// TIA Portal V17 export
// export: Created 2026-11-08T05:50:28.6935429Z, ExportSetting WithDefaults, DisplayName Totally Integrated Automation Portal, DisplayVersion V17, DisplayName TIA Portal Openness, DisplayVersion V17, DisplayName TIA Portal Version Control Interface, DisplayVersion V17, DisplayName STEP 7 Professional, DisplayVersion V17, DisplayName STEP 7 Safety, DisplayVersion V17, DisplayName WinCC Professional, DisplayVersion V17
FUNCTION_BLOCK "FB_Motor_Banderas"   // FB3, LAD
TITLE = Arranque y paro por BANDERAS (S/R)
{ S7_Optimized_Access := 'TRUE' }
VERSION : 0.1
// Estilo clásico: bandera de marcha con SET/RESET (paro dominante). Sin térmico se para; al recuperarse el térmico se puede volver a arrancar sin RESET.
// stored: AutoNumber true, IsIECCheckEnabled false, IsRetainMemResEnabled false, MemoryReserve 100, SetENOAutomatically false, UDAEnableTagReadback false
   VAR_INPUT
      Marcha : Bool;   // Orden de marcha (pulsador o HMI)
      Paro : Bool;   // Orden de paro: 1 = parar
      Termico_OK : Bool;   // 1 = relé térmico sin falla
      Reset : Bool;   // Reset de falla
   END_VAR
   VAR_OUTPUT
      Motor : Bool;   // Orden al contactor
      Piloto_Marcha : Bool;   // Piloto verde
      Piloto_Falla : Bool;   // Piloto rojo
      Estado : Int;   // 0 Reposo, 10 Marcha, 90 Falla
   END_VAR
   VAR
      B_Marcha : Bool;   // Bandera: motor en marcha
      B_Falla : Bool;   // Bandera: falla térmico
   END_VAR
BEGIN

REGION Network 1: SET bandera de marcha
   // Marcha sin paro y con térmico OK.
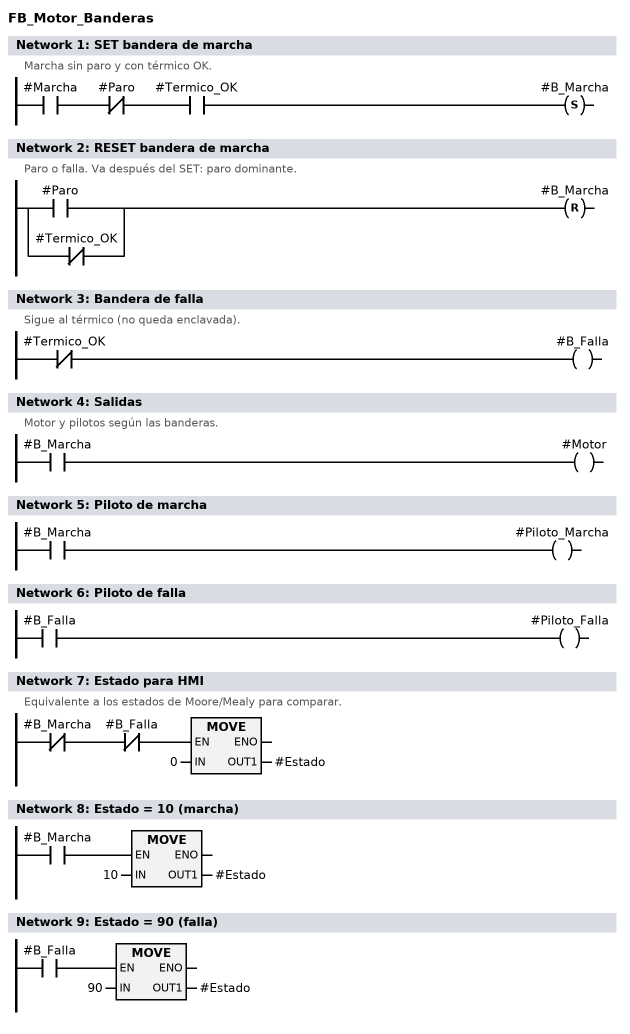
   RUNG wire#powerrail
      Contact( #Marcha )
      I_Contact( #Paro )
      Contact( #Termico_OK )
      S_Coil( #B_Marcha )
   END_RUNG
   // the same network as SCL:
   IF #Marcha AND NOT #Paro AND #Termico_OK THEN #B_Marcha := TRUE; END_IF;
END_REGION

REGION Network 2: RESET bandera de marcha
   // Paro o falla. Va después del SET: paro dominante.
   RUNG wire#powerrail
      Contact( #Paro )
      wire#w1
      R_Coil( #B_Marcha )
   END_RUNG
   RUNG wire#powerrail
      I_Contact( #Termico_OK )
   END_RUNG wire#w1
   // the same network as SCL:
   IF #Paro OR NOT #Termico_OK THEN #B_Marcha := FALSE; END_IF;
END_REGION

REGION Network 3: Bandera de falla
   // Sigue al térmico (no queda enclavada).
   RUNG wire#powerrail
      I_Contact( #Termico_OK )
      Coil( #B_Falla )
   END_RUNG
   // the same network as SCL:
   #B_Falla := NOT #Termico_OK;
END_REGION

REGION Network 4: Salidas
   // Motor y pilotos según las banderas.
   RUNG wire#powerrail
      Contact( #B_Marcha )
      Coil( #Motor )
   END_RUNG
   // the same network as SCL:
   #Motor := #B_Marcha;
END_REGION

REGION Network 5: Piloto de marcha
   RUNG wire#powerrail
      Contact( #B_Marcha )
      Coil( #Piloto_Marcha )
   END_RUNG
   // the same network as SCL:
   #Piloto_Marcha := #B_Marcha;
END_REGION

REGION Network 6: Piloto de falla
   RUNG wire#powerrail
      Contact( #B_Falla )
      Coil( #Piloto_Falla )
   END_RUNG
   // the same network as SCL:
   #Piloto_Falla := #B_Falla;
END_REGION

REGION Network 7: Estado para HMI
   // Equivalente a los estados de Moore/Mealy para comparar.
   RUNG wire#powerrail
      I_Contact( #B_Marcha )
      I_Contact( #B_Falla )
      { S7_GenerateENO := "TRUE" } Move(in := 0, out1 => #Estado)
   END_RUNG
   // the same network as SCL:
   IF NOT #B_Marcha AND NOT #B_Falla THEN #Estado := 0; END_IF;
END_REGION

REGION Network 8: Estado = 10 (marcha)
   RUNG wire#powerrail
      Contact( #B_Marcha )
      { S7_GenerateENO := "TRUE" } Move(in := 10, out1 => #Estado)
   END_RUNG
   // the same network as SCL:
   IF #B_Marcha THEN #Estado := 10; END_IF;
END_REGION

REGION Network 9: Estado = 90 (falla)
   RUNG wire#powerrail
      Contact( #B_Falla )
      { S7_GenerateENO := "TRUE" } Move(in := 90, out1 => #Estado)
   END_RUNG
   // the same network as SCL:
   IF #B_Falla THEN #Estado := 90; END_IF;
END_REGION
END_FUNCTION_BLOCK
